// TIA Portal project "OmronFQ2sensor30012026HardInterupt2IRT" (V17)

(* hardware
DEVICE "S7-1200 station_1"  S7-1200 Station
   slot 0: "Rack_0"  S7-1200 Rack  Rack  V1.0
   slot 1: "PLC_1"  CPU 1215C DC/DC/Rly  6ES7 215-1HG40-0XB0  V4.2
DEVICE "FQ2"  GSD.Device.PN
   slot 0: "Rack"  Rack  V1.0
   slot 0: "FQ2"  FQ2-XXX  FQ2-XXX  1.9.0
      slot 0: "FQ2-XXX"  FQ2-XXX  1.9.0
      slot 1: "Interface"  Interface
         slot 1: "Port 1"  Port 1
      slot 1: "Output Data_1"  Output Data  1.9.0
         slot 0: "Output Data"  Output Data  1.9.0
   slot 2: "Results Data - 32 items_1"  Results Data - 32 items  1.9.0
      slot 0: "Results Data - 32 items"  Results Data - 32 items  1.9.0
DEVICE "GSD device_1"  GSD.Device.PN
   slot 0: "Rack"  Rack  V1.0
   slot 0: "FQ22"  FQ2-XXX  FQ2-XXX  1.9.0
      slot 0: "FQ2-XXX"  FQ2-XXX  1.9.0
      slot 1: "Interface"  Interface
         slot 1: "Port 1"  Port 1
      slot 1: "Output Data_1"  Output Data  1.9.0
         slot 0: "Output Data"  Output Data  1.9.0
   slot 2: "Results Data - 32 items_1"  Results Data - 32 items  1.9.0
      slot 0: "Results Data - 32 items"  Results Data - 32 items  1.9.0
*)

// ===== PLC "PLC_1"  CPU 1215C DC/DC/Rly =====

VAR_GLOBAL   // PLC tag table "FQ2"
   "HWCurrentImpulseEncoder" AT %ID1000 : DInt;   // Значение счётчика энкодера в CPU
   "Input_Discret_Sensor_Product" AT %I0.7 : Bool;   // Входа наличия продукта
   "DOPusher" AT %Q0.0 : Bool;   // Выхода на отбраковщик
   "TemplVariable1ForFront" AT %M100.0 : Bool;   // Временая переменная для формирования фронта счёт продука
   "TempleVarible2ForFront" AT %M100.1 : Bool;   // Временая переменая для формирования фронта счёта брака
   "TempleVarible3ForFront" AT %M100.2 : Bool;
   "Tag_1" AT %M100.5 : Bool;
   "Tag_2" AT %M10.1 : Bool;
   "TempleVarible4ForFront" AT %M100.3 : Bool;
   "TempleVarible5ForFront" AT %M100.4 : Bool;
   "Tag_3" AT %M0.0 : Bool;
END_VAR

DATA_BLOCK "QueueProduct_1"   // DB1
{ S7_Optimized_Access := 'FALSE' }
VERSION : 0.1
   VAR
      StructQueue : Array[0..100] of Struct
         QueueAwaitingTrigerCam : Bool;   // Бит ожидания в очереди по камере
         QueueAwaitingRejection : Bool;   // Бит ожидания в очереди по отбраковке
         AwaitingDistanceCamera : Bool;   // Бит ожидание пройденой дистанции до камеры
         ActiveTrigerCam : Bool;   // Бит на измерение камеры
         AwaitingResultatMeasurement : Bool;   // Бит состояния ожидания ответа от камеры
         ResultMeasurementCamera : Bool;   // Результат полученый от камеры 0-ок 1-брак
         ResultRecieved : Bool;   // Результат получен
         RejectionOn : Bool;   // Активент отбраковщик
         CurrentImpulseEncodera : DInt;
      END_STRUCT;
   END_VAR
BEGIN
END_DATA_BLOCK

DATA_BLOCK "InputOutputCamer"   // DB2
{ S7_Optimized_Access := 'FALSE' }
VERSION : 0.1
   VAR
      InputFromCamera1 : Struct
         FLG : Bool;
         BUSY : Bool;
         Ready : Bool;
         "OR" : Bool;
         RUN : Bool;
         Resv : Bool;
         Resv_1 : Bool;
         Resv_2 : Bool;
         Resv_3 : Bool;
         Resv_4 : Bool;
         Resv_5 : Bool;
         Resv_6 : Bool;
         Resv_7 : Bool;
         Resv_8 : Bool;
         Resv_9 : Bool;
         Error : Bool;
         Gate : Bool;
         Resv_10 : Bool;
         Resv_11 : Bool;
         Resv_12 : Bool;
         Resv_13 : Bool;
         Resv_14 : Bool;
         Resv_15 : Bool;
         Resv_16 : Bool;
         Resv_17 : Bool;
         Resv_18 : Bool;
         Resv_19 : Bool;
         Resv_20 : Bool;
         Resv_21 : Bool;
         Resv_22 : Bool;
         Resv_23 : Bool;
         Resv_24 : Bool;
         CommandCode : Array[0..1] of Word;
         ResponseCode : Array[0..3] of Byte;
         ResponseData : Array[0..3] of Byte;
         OutputData1 : Array[0..3] of Byte;
         OutputData2 : Array[0..3] of Byte;
         OutputData3 : Array[0..3] of Byte;
         OutputData4 : Array[0..3] of Byte;
         OutputData5 : Array[0..3] of Byte;
         OutputData6 : Array[0..3] of Byte;
         OutputData7 : Array[0..3] of Byte;
         OutputData8 : Array[0..3] of Byte;
         OutputData9 : Array[0..3] of Byte;
         OutputData10 : Array[0..3] of Byte;
         OutputData11 : Array[0..3] of Byte;
         OutputData12 : Array[0..3] of Byte;
         OutputData13 : Array[0..3] of Byte;
         OutputData14 : Array[0..3] of Byte;
         OutputData15 : Array[0..3] of Byte;
         OutputData16 : Array[0..3] of Byte;
         OutputData17 : Array[0..3] of Byte;
         OutputData18 : Array[0..3] of Byte;
         OutputData19 : Array[0..3] of Byte;
         OutputData20 : Array[0..3] of Byte;
         OutputData21 : Array[0..3] of Byte;
         OutputData22 : Array[0..3] of Byte;
         OutputData23 : Array[0..3] of Byte;
         OutputData24 : Array[0..3] of Byte;
         OutputData25 : Array[0..3] of Byte;
         OutputData26 : Array[0..3] of Byte;
         OutputData27 : Array[0..3] of Byte;
         OutputData28 : Array[0..3] of Byte;
         OutputData29 : Array[0..3] of Byte;
         OutputData30 : Array[0..3] of Byte;
         OutputData31 : Array[0..3] of Byte;
         OutputData32 : Array[0..3] of Byte;
      END_STRUCT;
      OutputFromPLCtoCamera1 : Struct
         EXE : Bool;
         TRIG : Bool;
         Resv : Bool;
         Resv_1 : Bool;
         Resv_2 : Bool;
         Resv_3 : Bool;
         Resv_4 : Bool;
         Resv_5 : Bool;
         Resv_6 : Bool;
         Resv_7 : Bool;
         Resv_8 : Bool;
         Resv_9 : Bool;
         Resv_10 : Bool;
         Resv_11 : Bool;
         Resv_12 : Bool;
         ERCLR : Bool;
         DSA : Bool;
         Resv_13 : Bool;
         Resv_14 : Bool;
         Resv_15 : Bool;
         Resv_16 : Bool;
         Resv_17 : Bool;
         Resv_18 : Bool;
         Resv_19 : Bool;
         Resv_20 : Bool;
         Resv_21 : Bool;
         Resv_22 : Bool;
         Resv_23 : Bool;
         Resv_24 : Bool;
         Resv_25 : Bool;
         Resv_26 : Bool;
         Resv_27 : Bool;
         ComandCode : Array[0..1] of Word;
         ComandParameter : Array[0..3] of Byte;
         ComandParameter2 : Array[0..3] of Byte;
         ComandParameter3 : Array[0..3] of Byte;
      END_STRUCT;
      InputFromCamera2 : Struct
         FLG : Bool;
         BUSY : Bool;
         Ready : Bool;
         "OR" : Bool;
         RUN : Bool;
         Resv : Bool;
         Resv_1 : Bool;
         Resv_2 : Bool;
         Resv_3 : Bool;
         Resv_4 : Bool;
         Resv_5 : Bool;
         Resv_6 : Bool;
         Resv_7 : Bool;
         Resv_8 : Bool;
         Resv_9 : Bool;
         Error : Bool;
         Gate : Bool;
         Resv_10 : Bool;
         Resv_11 : Bool;
         Resv_12 : Bool;
         Resv_13 : Bool;
         Resv_14 : Bool;
         Resv_15 : Bool;
         Resv_16 : Bool;
         Resv_17 : Bool;
         Resv_18 : Bool;
         Resv_19 : Bool;
         Resv_20 : Bool;
         Resv_21 : Bool;
         Resv_22 : Bool;
         Resv_23 : Bool;
         Resv_24 : Bool;
         CommandCode : Array[0..1] of Word;
         ResponseCode : Array[0..3] of Byte;
         ResponseData : Array[0..3] of Byte;
         OutputData1 : Array[0..3] of Byte;
         OutputData2 : Array[0..3] of Byte;
         OutputData3 : Array[0..3] of Byte;
         OutputData4 : Array[0..3] of Byte;
         OutputData5 : Array[0..3] of Byte;
         OutputData6 : Array[0..3] of Byte;
         OutputData7 : Array[0..3] of Byte;
         OutputData8 : Array[0..3] of Byte;
         OutputData9 : Array[0..3] of Byte;
         OutputData10 : Array[0..3] of Byte;
         OutputData11 : Array[0..3] of Byte;
         OutputData12 : Array[0..3] of Byte;
         OutputData13 : Array[0..3] of Byte;
         OutputData14 : Array[0..3] of Byte;
         OutputData15 : Array[0..3] of Byte;
         OutputData16 : Array[0..3] of Byte;
         OutputData17 : Array[0..3] of Byte;
         OutputData18 : Array[0..3] of Byte;
         OutputData19 : Array[0..3] of Byte;
         OutputData20 : Array[0..3] of Byte;
         OutputData21 : Array[0..3] of Byte;
         OutputData22 : Array[0..3] of Byte;
         OutputData23 : Array[0..3] of Byte;
         OutputData24 : Array[0..3] of Byte;
         OutputData25 : Array[0..3] of Byte;
         OutputData26 : Array[0..3] of Byte;
         OutputData27 : Array[0..3] of Byte;
         OutputData28 : Array[0..3] of Byte;
         OutputData29 : Array[0..3] of Byte;
         OutputData30 : Array[0..3] of Byte;
         OutputData31 : Array[0..3] of Byte;
         OutputData32 : Array[0..3] of Byte;
      END_STRUCT;
      OutputFromPLCtoCamera2 : Struct
         EXE : Bool;
         TRIG : Bool;
         Resv : Bool;
         Resv_1 : Bool;
         Resv_2 : Bool;
         Resv_3 : Bool;
         Resv_4 : Bool;
         Resv_5 : Bool;
         Resv_6 : Bool;
         Resv_7 : Bool;
         Resv_8 : Bool;
         Resv_9 : Bool;
         Resv_10 : Bool;
         Resv_11 : Bool;
         Resv_12 : Bool;
         ERCLR : Bool;
         DSA : Bool;
         Resv_13 : Bool;
         Resv_14 : Bool;
         Resv_15 : Bool;
         Resv_16 : Bool;
         Resv_17 : Bool;
         Resv_18 : Bool;
         Resv_19 : Bool;
         Resv_20 : Bool;
         Resv_21 : Bool;
         Resv_22 : Bool;
         Resv_23 : Bool;
         Resv_24 : Bool;
         Resv_25 : Bool;
         Resv_26 : Bool;
         Resv_27 : Bool;
         ComandCode : Array[0..1] of Word;
         ComandParameter : Array[0..3] of Byte;
         ComandParameter2 : Array[0..3] of Byte;
         ComandParameter3 : Array[0..3] of Byte;
      END_STRUCT;
   END_VAR
BEGIN
   InputFromCamera1.CommandCode[0] := 16#0;
   InputFromCamera2.CommandCode[0] := 16#0;
END_DATA_BLOCK

DATA_BLOCK "AuxaluryBlockProcesseComandeCamera"   // DB3
{ S7_Optimized_Access := 'FALSE' }
VERSION : 0.1
   VAR
      RequestComandeFromPlcToCamera_1 : Bool;   // Бит начала запроса выполнения команды с плк на камеру
      RequestConfirmComandeFromPLCtoCamera_1 : Bool;   // Бит подтверждения что запрос команды отправлен
      RequestComandeFromPlcToCamera_2 : Bool;
      RequestConfirmComandeFromPLCtoCamera_2 : Bool;
      Camera1ChangeSceneOk : Bool;
      Camera2ChangeSceneOk : Bool;
      QuitRejectCam1 : Bool;   // Отбраковка по камере 1
      QuitRejectCam2 : Bool;   // Отбраковка по камере 2
      RequestChangeSceneCamera1 : Bool;   // Дополнительный бить для обработки переключения рецецтпа камеры 1
      RequestChangeSceneCamera2 : Bool;   // Дополнительный бить для обработки переключения рецецтпа камеры 2
   END_VAR
BEGIN
END_DATA_BLOCK

DATA_BLOCK "QueueProduct_2"   // DB4
{ S7_Optimized_Access := 'TRUE' }
VERSION : 0.1
   VAR
      StructQueue : Array[0..100] of Struct
         QueueAwaitingTrigerCam : Bool;   // Бит ожидания в очереди по камере
         QueueAwaitingRejection : Bool;   // Бит ожидания в очереди по отбраковке
         AwaitingDistanceCamera : Bool;   // Бит ожидание пройденой дистанции до камеры
         ActiveTrigerCam : Bool;   // Бит на измерение камеры
         AwaitingResultatMeasurement : Bool;   // Бит состояния ожидания ответа от камеры
         ResultMeasurementCamera : Bool;   // Результат полученый от камеры 0-ок 1-брак
         ResultRecieved : Bool;   // Результат получен
         RejectionOn : Bool;   // Активент отбраковщик
         CurrentImpulseEncodera : DInt;
      END_STRUCT;
   END_VAR
BEGIN
END_DATA_BLOCK

DATA_BLOCK "DataBlockHMI"   // DB5
{ S7_Optimized_Access := 'FALSE' }
VERSION : 0.1
   VAR
      CountProduct : UDInt;   // Кол-во продукта прошедшего отбраковщик
      CountRejection : UDInt;   // Кол-во отбракованного
      NumberSceneRequest : Byte;   // Запрос номера сценария в камере
      Buttons : Struct
         ButtonChangeRecipe : Bool;   // Кнопка запрос на изменение рецепта(сцены)камеры от оператора
         ButtonWorkRestrictionPusher : Bool;   // Кнопка запрета работы пушера отбраковщика
         ButtonLoadFromActualInList : Bool;
         ButtonWorkOffCam1 : Bool;   // Камера 1 не обрабатывает очередь продукта
         ButtonWorkOffCam2 : Bool;   // Камера 2 не обрабатывает очередь продукта
         Button5 : Bool;
         Button6 : Bool;
         Button7 : Bool;
      END_STRUCT;
      AuxilaryBit : Array[0..7] of Bool;
      Recipe : Array[0..32] of Struct
         CountImpTrigerCamera1 : DInt;   // Количество импульсов для сработки камеры
         CountImpForRegection1 : DInt;   // Количество импульсов для отбраковки
         CountImpForResetRegectio1 : DInt;   // Количество импульсов для длительности отбраковки
         NumberRecipeScene : Byte;   // Номер сценария в камере
         HighMM : Int;   // высота в милиметрах
         OverhangValue : Int;   // величина вылета в милиметрах
         CountImpTrigerCamera2 : DInt;
         CountImpForRegection2 : DInt;
      END_STRUCT;
      CountRejectionCam1 : UDInt;   // Количество отбраковоаного по камере 1
      CountRejectionCam2 : UDInt;   // Количество отбракованого по камере 2
   END_VAR
BEGIN
   Recipe[0].CountImpTrigerCamera1 := 335;
   Recipe[0].CountImpForRegection1 := 455;
   Recipe[0].CountImpForResetRegectio1 := 25;
   Recipe[0].NumberRecipeScene := 0;
   Recipe[1].CountImpTrigerCamera1 := 335;
   Recipe[1].CountImpForRegection1 := 455;
   Recipe[1].CountImpForResetRegectio1 := 25;
   Recipe[1].NumberRecipeScene := 0;
   Recipe[2].CountImpTrigerCamera1 := 335;
   Recipe[2].CountImpForRegection1 := 455;
   Recipe[2].CountImpForResetRegectio1 := 25;
   Recipe[2].NumberRecipeScene := 1;
   Recipe[3].CountImpTrigerCamera1 := 335;
   Recipe[3].CountImpForRegection1 := 455;
   Recipe[3].CountImpForResetRegectio1 := 25;
   Recipe[3].NumberRecipeScene := 2;
   Recipe[4].CountImpTrigerCamera1 := 335;
   Recipe[4].CountImpForRegection1 := 455;
   Recipe[4].CountImpForResetRegectio1 := 25;
   Recipe[4].NumberRecipeScene := 3;
   Recipe[5].CountImpTrigerCamera1 := 335;
   Recipe[5].CountImpForRegection1 := 455;
   Recipe[5].CountImpForResetRegectio1 := 25;
   Recipe[5].NumberRecipeScene := 4;
   Recipe[6].CountImpTrigerCamera1 := 335;
   Recipe[6].CountImpForRegection1 := 455;
   Recipe[6].CountImpForResetRegectio1 := 25;
   Recipe[6].NumberRecipeScene := 5;
   Recipe[7].CountImpTrigerCamera1 := 335;
   Recipe[7].CountImpForRegection1 := 455;
   Recipe[7].CountImpForResetRegectio1 := 25;
   Recipe[7].NumberRecipeScene := 6;
   Recipe[8].CountImpTrigerCamera1 := 335;
   Recipe[8].CountImpForRegection1 := 455;
   Recipe[8].CountImpForResetRegectio1 := 25;
   Recipe[8].NumberRecipeScene := 7;
   Recipe[9].CountImpTrigerCamera1 := 335;
   Recipe[9].CountImpForRegection1 := 455;
   Recipe[9].CountImpForResetRegectio1 := 25;
   Recipe[9].NumberRecipeScene := 8;
   Recipe[10].CountImpTrigerCamera1 := 335;
   Recipe[10].CountImpForRegection1 := 455;
   Recipe[10].CountImpForResetRegectio1 := 25;
   Recipe[10].NumberRecipeScene := 9;
   Recipe[11].CountImpTrigerCamera1 := 335;
   Recipe[11].CountImpForRegection1 := 455;
   Recipe[11].CountImpForResetRegectio1 := 25;
   Recipe[11].NumberRecipeScene := 10;
   Recipe[12].CountImpTrigerCamera1 := 335;
   Recipe[12].CountImpForRegection1 := 455;
   Recipe[12].CountImpForResetRegectio1 := 25;
   Recipe[12].NumberRecipeScene := 11;
   Recipe[13].CountImpTrigerCamera1 := 335;
   Recipe[13].CountImpForRegection1 := 455;
   Recipe[13].CountImpForResetRegectio1 := 25;
   Recipe[13].NumberRecipeScene := 12;
   Recipe[14].CountImpTrigerCamera1 := 335;
   Recipe[14].CountImpForRegection1 := 455;
   Recipe[14].CountImpForResetRegectio1 := 25;
   Recipe[14].NumberRecipeScene := 13;
   Recipe[15].CountImpTrigerCamera1 := 335;
   Recipe[15].CountImpForRegection1 := 455;
   Recipe[15].CountImpForResetRegectio1 := 25;
   Recipe[15].NumberRecipeScene := 14;
   Recipe[16].CountImpTrigerCamera1 := 335;
   Recipe[16].CountImpForRegection1 := 455;
   Recipe[16].CountImpForResetRegectio1 := 25;
   Recipe[16].NumberRecipeScene := 15;
   Recipe[17].CountImpTrigerCamera1 := 335;
   Recipe[17].CountImpForRegection1 := 455;
   Recipe[17].CountImpForResetRegectio1 := 25;
   Recipe[17].NumberRecipeScene := 16;
   Recipe[18].CountImpTrigerCamera1 := 335;
   Recipe[18].CountImpForRegection1 := 455;
   Recipe[18].CountImpForResetRegectio1 := 25;
   Recipe[18].NumberRecipeScene := 17;
   Recipe[19].CountImpTrigerCamera1 := 335;
   Recipe[19].CountImpForRegection1 := 455;
   Recipe[19].CountImpForResetRegectio1 := 25;
   Recipe[19].NumberRecipeScene := 18;
   Recipe[20].CountImpTrigerCamera1 := 335;
   Recipe[20].CountImpForRegection1 := 455;
   Recipe[20].CountImpForResetRegectio1 := 25;
   Recipe[20].NumberRecipeScene := 19;
   Recipe[21].CountImpTrigerCamera1 := 335;
   Recipe[21].CountImpForRegection1 := 455;
   Recipe[21].CountImpForResetRegectio1 := 25;
   Recipe[21].NumberRecipeScene := 20;
   Recipe[22].CountImpTrigerCamera1 := 335;
   Recipe[22].CountImpForRegection1 := 455;
   Recipe[22].CountImpForResetRegectio1 := 25;
   Recipe[22].NumberRecipeScene := 21;
   Recipe[23].CountImpTrigerCamera1 := 335;
   Recipe[23].CountImpForRegection1 := 455;
   Recipe[23].CountImpForResetRegectio1 := 25;
   Recipe[23].NumberRecipeScene := 22;
   Recipe[24].CountImpTrigerCamera1 := 335;
   Recipe[24].CountImpForRegection1 := 455;
   Recipe[24].CountImpForResetRegectio1 := 25;
   Recipe[24].NumberRecipeScene := 23;
   Recipe[25].CountImpTrigerCamera1 := 335;
   Recipe[25].CountImpForRegection1 := 455;
   Recipe[25].CountImpForResetRegectio1 := 25;
   Recipe[25].NumberRecipeScene := 24;
   Recipe[26].CountImpTrigerCamera1 := 335;
   Recipe[26].CountImpForRegection1 := 455;
   Recipe[26].CountImpForResetRegectio1 := 25;
   Recipe[26].NumberRecipeScene := 25;
   Recipe[27].CountImpTrigerCamera1 := 335;
   Recipe[27].CountImpForRegection1 := 455;
   Recipe[27].CountImpForResetRegectio1 := 25;
   Recipe[27].NumberRecipeScene := 26;
   Recipe[28].CountImpTrigerCamera1 := 335;
   Recipe[28].CountImpForRegection1 := 455;
   Recipe[28].CountImpForResetRegectio1 := 25;
   Recipe[28].NumberRecipeScene := 27;
   Recipe[29].CountImpTrigerCamera1 := 335;
   Recipe[29].CountImpForRegection1 := 455;
   Recipe[29].CountImpForResetRegectio1 := 25;
   Recipe[29].NumberRecipeScene := 28;
   Recipe[30].CountImpTrigerCamera1 := 335;
   Recipe[30].CountImpForRegection1 := 455;
   Recipe[30].CountImpForResetRegectio1 := 25;
   Recipe[30].NumberRecipeScene := 29;
   Recipe[31].CountImpTrigerCamera1 := 335;
   Recipe[31].CountImpForRegection1 := 455;
   Recipe[31].CountImpForResetRegectio1 := 25;
   Recipe[31].NumberRecipeScene := 30;
   Recipe[32].CountImpTrigerCamera1 := 335;
   Recipe[32].CountImpForRegection1 := 455;
   Recipe[32].CountImpForResetRegectio1 := 25;
   Recipe[32].NumberRecipeScene := 31;
   // AuxilaryBit[0] : Бит для подсчёта брака cam1
   // Recipe[0] : Действующей рецепт(сценарий)
   // Recipe[1] : Сценарий 0
   // Recipe[2] : Сценарий 1
   // Recipe[3] : Сценарий 2
   // Recipe[4] : Сценарий 3
   // Recipe[5] : Сценарий 4
   // Recipe[6] : Сценарий 5
   // Recipe[7] : Сценарий 6
   // Recipe[8] : Сценарий 7
   // Recipe[9] : Сценарий 8
   // Recipe[10] : Сценарий 9
   // AuxilaryBit[1] : Бит для подсчёта брака сam2
END_DATA_BLOCK

FUNCTION "QueueCreate" : Void   // FC3, SCL
{ S7_Optimized_Access := 'FALSE' }
VERSION : 0.1
   VAR_TEMP
      i1 : Int;
      i2 : Int;
      d : Int;
   END_VAR
BEGIN
   //Добовляем в очередь продукт

       FOR #i1 := 0 TO 20 DO
           // Statement section FOR
           IF NOT "QueueProduct_1".StructQueue[#i1].QueueAwaitingRejection THEN
               IF NOT "DataBlockHMI".Buttons.ButtonWorkOffCam1 THEN //условие чтоб камеру выключить не обрабоатывать ничего
                   "QueueProduct_1".StructQueue[#i1].QueueAwaitingTrigerCam := TRUE;
                   "QueueProduct_1".StructQueue[#i1].QueueAwaitingRejection := TRUE;
               END_IF;

               EXIT;
           END_IF;
       END_FOR;
       FOR #i2 := 0 TO 20 DO
           // Statement section FOR
           IF NOT "QueueProduct_2".StructQueue[#i2].QueueAwaitingRejection THEN
               IF NOT "DataBlockHMI".Buttons.ButtonWorkOffCam2 THEN
                   "QueueProduct_2".StructQueue[#i2].QueueAwaitingTrigerCam := TRUE;
                   "QueueProduct_2".StructQueue[#i2].QueueAwaitingRejection := TRUE;
               END_IF;
               EXIT;
           END_IF;
       END_FOR;

   "DataBlockHMI".CountProduct := UDINT#1 + "DataBlockHMI".CountProduct;

   IF NOT "DataBlockHMI".Buttons.ButtonWorkOffCam1 THEN
       "ProcessingQueue1"(NumberQueue := #i1); //Обрабатываем только что добавленую очередь
   END_IF;
   IF NOT "DataBlockHMI".Buttons.ButtonWorkOffCam2 THEN
       "ProcessingQueue2"(NumberQueue := #i2);
   END_IF;
END_FUNCTION

FUNCTION "ProcessingQueue1" : Void   // FC4, SCL
{ S7_Optimized_Access := 'TRUE' }
VERSION : 0.1
   VAR_INPUT
      NumberQueue : Int;
   END_VAR
BEGIN
   IF  "QueueProduct_1".StructQueue[#NumberQueue].QueueAwaitingRejection THEN
       // Statement section IF


       //Создание запроса в очереди на тригер камеры, запоминаем текущие положение продукта
       IF "QueueProduct_1".StructQueue[#NumberQueue].QueueAwaitingTrigerCam &
           "QueueProduct_1".StructQueue[#NumberQueue].QueueAwaitingRejection THEN

           "QueueProduct_1".StructQueue[#NumberQueue].CurrentImpulseEncodera := "HWCurrentImpulseEncoder":P;
           "QueueProduct_1".StructQueue[#NumberQueue].QueueAwaitingTrigerCam := False;
           "QueueProduct_1".StructQueue[#NumberQueue].AwaitingDistanceCamera := True;
           RETURN;
       END_IF;
       //Выходим из проверки пока продукт не доехал до камеры, оптимизация чтоб не пробегать всю функцию
       IF "QueueProduct_1".StructQueue[#NumberQueue].CurrentImpulseEncodera +"DataBlockHMI".Recipe[0].CountImpTrigerCamera1(*Recip[0] прният как действующей рецепт*) >"HWCurrentImpulseEncoder":P THEN
           RETURN;
       END_IF;    
           //По прохождению дистанции взводим бит для работы камеры, снимаем бит ожидания 
       IF "QueueProduct_1".StructQueue[#NumberQueue].AwaitingDistanceCamera
           &"QueueProduct_1".StructQueue[#NumberQueue].CurrentImpulseEncodera + "DataBlockHMI".Recipe[0].CountImpTrigerCamera1(*Recip[0] прният как действующей рецепт*) <="HWCurrentImpulseEncoder":P
            & NOT "InputOutputCamer".InputFromCamera1.BUSY THEN

           "QueueProduct_1".StructQueue[#NumberQueue].ActiveTrigerCam := true;
           "InputOutputCamer".OutputFromPLCtoCamera1.TRIG := true;
           "QueueProduct_1".StructQueue[#NumberQueue].AwaitingDistanceCamera := False;
           RETURN;
       END_IF;

       //На период обработки камеры снимаем бит работы камеры, взводим бит ожидание ответа от камеры
       IF "QueueProduct_1".StructQueue[#NumberQueue].ActiveTrigerCam & "InputOutputCamer".InputFromCamera1.BUSY THEN

           "QueueProduct_1".StructQueue[#NumberQueue].ActiveTrigerCam := False;
           "InputOutputCamer".OutputFromPLCtoCamera1.TRIG := false;
           "QueueProduct_1".StructQueue[#NumberQueue].AwaitingResultatMeasurement := True;
           RETURN;
       END_IF;

       //Ожидание получение ответа от камеры, фиксируем что ответ был
       IF "QueueProduct_1".StructQueue[#NumberQueue].AwaitingResultatMeasurement & NOT "InputOutputCamer".InputFromCamera1.BUSY
       THEN

           "QueueProduct_1".StructQueue[#NumberQueue].ResultMeasurementCamera := "InputOutputCamer".InputFromCamera1."OR";
           "QueueProduct_1".StructQueue[#NumberQueue].ResultRecieved := True;
           "QueueProduct_1".StructQueue[#NumberQueue].AwaitingResultatMeasurement := FALSE;

       END_IF;

       //Обработка полученого ответа от камеры(бракуем или нет).
       //Если не бракуем, освобождаем очередь, Если бракуем то взводим бит браковки и освобождаем очередь после снятия сигнала с пушера
       IF "QueueProduct_1".StructQueue[#NumberQueue].ResultRecieved & "QueueProduct_1".StructQueue[#NumberQueue].ResultMeasurementCamera
           & ("QueueProduct_1".StructQueue[#NumberQueue].CurrentImpulseEncodera + "DataBlockHMI".Recipe[0].CountImpTrigerCamera1
           + "DataBlockHMI".Recipe[0].CountImpForRegection1 <= "HWCurrentImpulseEncoder":P) THEN //условия для старта отбраковки

           "AuxaluryBlockProcesseComandeCamera".QuitRejectCam1 := true;
           "DataBlockHMI".AuxilaryBit[0] := TRUE;
           "QueueProduct_1".StructQueue[#NumberQueue].RejectionOn := true;
           "QueueProduct_1".StructQueue[#NumberQueue].ResultRecieved := FALSE;

       ELSIF "QueueProduct_1".StructQueue[#NumberQueue].ResultRecieved & NOT "QueueProduct_1".StructQueue[#NumberQueue].ResultMeasurementCamera THEN

           "QueueProduct_1".StructQueue[#NumberQueue] := "QueueProduct_1".StructQueue[100];

       END_IF;

       //Cнимаем выход отбраковки и скидываем очередь
       IF "QueueProduct_1".StructQueue[#NumberQueue].RejectionOn & ("QueueProduct_1".StructQueue[#NumberQueue].CurrentImpulseEncodera + "DataBlockHMI".Recipe[0].CountImpTrigerCamera1
           + "DataBlockHMI".Recipe[0].CountImpForRegection1 +"DataBlockHMI".Recipe[0].CountImpForResetRegectio1 <="HWCurrentImpulseEncoder":P) THEN

           "AuxaluryBlockProcesseComandeCamera".QuitRejectCam1 := false;
           "DataBlockHMI".AuxilaryBit[0] := FALSE;
           "QueueProduct_1".StructQueue[#NumberQueue] := "QueueProduct_1".StructQueue[100];

       END_IF;

       IF "DataBlockHMI".Buttons.ButtonWorkRestrictionPusher THEN
           "AuxaluryBlockProcesseComandeCamera".QuitRejectCam1 := FALSE;

       END_IF;


   END_IF;
END_FUNCTION

FUNCTION "ChangeSceneOnCameraFQ2" : Void   // FC6, SCL
{ S7_Optimized_Access := 'FALSE' }
VERSION : 0.1
   VAR_INPUT
      NumberScene : Byte;
   END_VAR
   VAR_IN_OUT
      RequestChangeScene : Bool;
   END_VAR
BEGIN
   //Запроc смены рецепта или есть ожидание от прошлого выполняем
   //условия обработки смены сценария, здесь создаём защиту от зацикливания
   //посредсвом проверки прошлый запрос прошёл успешно и ждём вторую камеру

   IF #RequestChangeScene AND NOT "AuxaluryBlockProcesseComandeCamera".RequestChangeSceneCamera1 AND NOT "AuxaluryBlockProcesseComandeCamera".Camera1ChangeSceneOk THEN
          "AuxaluryBlockProcesseComandeCamera".RequestChangeSceneCamera1 := TRUE;
      END_IF;

   IF #RequestChangeScene AND NOT "AuxaluryBlockProcesseComandeCamera".RequestChangeSceneCamera2 AND NOT "AuxaluryBlockProcesseComandeCamera".Camera2ChangeSceneOk THEN
         "AuxaluryBlockProcesseComandeCamera".RequestChangeSceneCamera2 := TRUE;
   END_IF;


   // Команда на камеру1 для выполнения переключения сценария проверки и номер сценария
      IF "AuxaluryBlockProcesseComandeCamera".RequestChangeSceneCamera1 AND NOT "InputOutputCamer".InputFromCamera1.BUSY
          AND NOT "AuxaluryBlockProcesseComandeCamera".Camera1ChangeSceneOk THEN


         "InputOutputCamer".OutputFromPLCtoCamera1.ComandCode[0] := 16#30;
         "InputOutputCamer".OutputFromPLCtoCamera1.ComandCode[1] := 16#1000;
         "InputOutputCamer".OutputFromPLCtoCamera1.ComandParameter[3] := #NumberScene;
         "AuxaluryBlockProcesseComandeCamera".RequestConfirmComandeFromPLCtoCamera_1 := TRUE;
         "InputOutputCamer".OutputFromPLCtoCamera1.EXE := TRUE;

     END_IF;

   // Команда на камеру2 для выполнения переключения сценария проверки и номер сценария
     IF "AuxaluryBlockProcesseComandeCamera".RequestChangeSceneCamera2 AND NOT "InputOutputCamer".InputFromCamera2.BUSY
         AND NOT "AuxaluryBlockProcesseComandeCamera".Camera2ChangeSceneOk THEN


         "InputOutputCamer".OutputFromPLCtoCamera2.ComandCode[0] := 16#30;
         "InputOutputCamer".OutputFromPLCtoCamera2.ComandCode[1] := 16#1000;
         "InputOutputCamer".OutputFromPLCtoCamera2.ComandParameter[3] := #NumberScene;
         "AuxaluryBlockProcesseComandeCamera".RequestConfirmComandeFromPLCtoCamera_2 := TRUE;
         "InputOutputCamer".OutputFromPLCtoCamera2.EXE := TRUE;

     END_IF;

       // После послания запроса ожидаем возвращени выполнения подтверждения от камеры 1, что всё выполнено и сбрасываем биты и команды.
     IF "AuxaluryBlockProcesseComandeCamera".RequestConfirmComandeFromPLCtoCamera_1
         AND "InputOutputCamer".InputFromCamera1.BUSY
         AND "InputOutputCamer".InputFromCamera1.FLG AND NOT "AuxaluryBlockProcesseComandeCamera".Camera1ChangeSceneOk THEN

         //#RequestChangeScene := FALSE;
         "AuxaluryBlockProcesseComandeCamera".RequestConfirmComandeFromPLCtoCamera_1 := FALSE;
         "InputOutputCamer".OutputFromPLCtoCamera1.EXE := False;
         "InputOutputCamer".OutputFromPLCtoCamera1.ComandCode[0] := 16#0;
         "InputOutputCamer".OutputFromPLCtoCamera1.ComandCode[1] := 16#0;
         "InputOutputCamer".OutputFromPLCtoCamera1.ComandParameter[3] := 0;
         IF "InputOutputCamer".InputFromCamera1.ResponseCode[0] = 0
             AND
             "InputOutputCamer".InputFromCamera1.ResponseCode[1] = 0
             AND
             "InputOutputCamer".InputFromCamera1.ResponseCode[2] = 0
             AND
             "InputOutputCamer".InputFromCamera1.ResponseCode[3] = 0
         THEN
             "AuxaluryBlockProcesseComandeCamera".Camera1ChangeSceneOk := TRUE;
         END_IF;
         //#RequestChangeScene := False;
     END_IF;

    // После послания запроса ожидаем возвращени выполнения подтверждения от камеры 2, что всё выполнено и сбрасываем биты и команды.
     IF "AuxaluryBlockProcesseComandeCamera".RequestConfirmComandeFromPLCtoCamera_2
         AND "InputOutputCamer".InputFromCamera2.BUSY
         AND "InputOutputCamer".InputFromCamera2.FLG AND NOT "AuxaluryBlockProcesseComandeCamera".Camera2ChangeSceneOk THEN

         //#RequestChangeScene := FALSE;
         "AuxaluryBlockProcesseComandeCamera".RequestConfirmComandeFromPLCtoCamera_2 := FALSE;
         "InputOutputCamer".OutputFromPLCtoCamera2.EXE := False;
         "InputOutputCamer".OutputFromPLCtoCamera2.ComandCode[0] := 16#0;
         "InputOutputCamer".OutputFromPLCtoCamera2.ComandCode[1] := 16#0;
         "InputOutputCamer".OutputFromPLCtoCamera2.ComandParameter[3] := 0;
         IF "InputOutputCamer".InputFromCamera2.ResponseCode[0] = 0
             AND
             "InputOutputCamer".InputFromCamera2.ResponseCode[1] = 0
             AND
             "InputOutputCamer".InputFromCamera2.ResponseCode[2] = 0
             AND
             "InputOutputCamer".InputFromCamera2.ResponseCode[3] = 0
         THEN
             "AuxaluryBlockProcesseComandeCamera".Camera2ChangeSceneOk:=TRUE;
         END_IF;
         //#RequestChangeScene := False;
     END_IF;
     (* IF "AuxaluryBlockProcesseComandeCamera".Camera1ChangeSceneOk  THEN
         "RecipeFromListToActual"(#NumberScene);
         //"AuxaluryBlockProcesseComandeCamera".Camera2ChangeSceneOk := FALSE;
         "AuxaluryBlockProcesseComandeCamera".Camera1ChangeSceneOk := FALSE;

     END_IF;

     IF "AuxaluryBlockProcesseComandeCamera".Camera2ChangeSceneOk THEN
         "RecipeFromListToActual"(#NumberScene);
         "AuxaluryBlockProcesseComandeCamera".Camera2ChangeSceneOk := FALSE;
         //"AuxaluryBlockProcesseComandeCamera".Camera1ChangeSceneOk := FALSE;

     END_IF; *)
     //Cнимаеме повторение запросов
     IF "AuxaluryBlockProcesseComandeCamera".Camera1ChangeSceneOk AND "AuxaluryBlockProcesseComandeCamera".RequestChangeSceneCamera1 THEN

         "AuxaluryBlockProcesseComandeCamera".RequestChangeSceneCamera1 := FALSE;

     END_IF;

     IF "AuxaluryBlockProcesseComandeCamera".Camera2ChangeSceneOk AND "AuxaluryBlockProcesseComandeCamera".RequestChangeSceneCamera2 THEN
         "AuxaluryBlockProcesseComandeCamera".RequestChangeSceneCamera1 := FALSE;
     END_IF;

     //Перенос рецепта из памяти в актуальный работающий сброс битов
     IF "AuxaluryBlockProcesseComandeCamera".Camera1ChangeSceneOk AND "AuxaluryBlockProcesseComandeCamera".Camera2ChangeSceneOk THEN
         "RecipeFromListToActual"(#NumberScene);
         "AuxaluryBlockProcesseComandeCamera".Camera1ChangeSceneOk := FALSE;
         "AuxaluryBlockProcesseComandeCamera".Camera2ChangeSceneOk := FALSE;
         #RequestChangeScene := FALSE;

     END_IF;
END_FUNCTION

FUNCTION "RecipeFromListToActual" : Void   // FC7, SCL
{ S7_Optimized_Access := 'TRUE' }
VERSION : 0.1
   VAR_INPUT
      InputNumber : Byte;   // Указание какой рецепт загружаем в актуальный
   END_VAR
   VAR_TEMP
      i : Int;   // временая переменая для прогона
   END_VAR
BEGIN

   FOR  #i:= 1 TO 32 DO

       IF "DataBlockHMI".Recipe[#i].NumberRecipeScene = #InputNumber THEN

           "DataBlockHMI".Recipe[0] := "DataBlockHMI".Recipe[#i];
           EXIT;
       END_IF;


       END_FOR;
END_FUNCTION

FUNCTION "RecipFromActualToList" : Void   // FC8, SCL
{ S7_Optimized_Access := 'TRUE' }
VERSION : 0.1
   VAR_INPUT
      InputNumber : Byte;
   END_VAR
   VAR_TEMP
      i : Int;
   END_VAR
BEGIN
   FOR #i := 1 TO 32 DO

       IF "DataBlockHMI".Recipe[#i].NumberRecipeScene = #InputNumber THEN

           "DataBlockHMI".Recipe[#i] := "DataBlockHMI".Recipe[0];
           EXIT;
       END_IF;


   END_FOR;
END_FUNCTION

FUNCTION "ProcessingQueue2" : Void   // FC9, SCL
{ S7_Optimized_Access := 'TRUE' }
VERSION : 0.1
   VAR_INPUT
      NumberQueue : Int;
   END_VAR
BEGIN
   IF "QueueProduct_2".StructQueue[#NumberQueue].QueueAwaitingRejection THEN
       // Statement section IF


       //Создание запроса в очереди на тригер камеры, запоминаем текущие положение продукта
       IF "QueueProduct_2".StructQueue[#NumberQueue].QueueAwaitingTrigerCam &
           "QueueProduct_2".StructQueue[#NumberQueue].QueueAwaitingRejection THEN

           "QueueProduct_2".StructQueue[#NumberQueue].CurrentImpulseEncodera := "HWCurrentImpulseEncoder":P;
           "QueueProduct_2".StructQueue[#NumberQueue].QueueAwaitingTrigerCam := False;
           "QueueProduct_2".StructQueue[#NumberQueue].AwaitingDistanceCamera := True;
           RETURN;
       END_IF;
       //Выходим из проверки пока продукт не доехал до камеры, оптимизация чтоб не пробегать всю функцию
       IF "QueueProduct_2".StructQueue[#NumberQueue].CurrentImpulseEncodera + "DataBlockHMI".Recipe[0].CountImpTrigerCamera2 > "HWCurrentImpulseEncoder":P THEN
           RETURN;
       END_IF;
       //По прохождению дистанции взводим бит для работы камеры, снимаем бит ожидания 
       IF  "QueueProduct_2".StructQueue[#NumberQueue].AwaitingDistanceCamera
           & "QueueProduct_2".StructQueue[#NumberQueue].CurrentImpulseEncodera + "DataBlockHMI".Recipe[0].CountImpTrigerCamera2<= "HWCurrentImpulseEncoder":P
           &  NOT "InputOutputCamer".InputFromCamera2.BUSY THEN

           "QueueProduct_2".StructQueue[#NumberQueue].ActiveTrigerCam := true;
           "InputOutputCamer".OutputFromPLCtoCamera2.TRIG := true;
           "QueueProduct_2".StructQueue[#NumberQueue].AwaitingDistanceCamera := False;
           RETURN;
       END_IF;

       //На период обработки камеры снимаем бит работы камеры, взводим бит ожидание ответа от камеры
       IF "QueueProduct_2".StructQueue[#NumberQueue].ActiveTrigerCam & "InputOutputCamer".InputFromCamera2.BUSY THEN

           "QueueProduct_2".StructQueue[#NumberQueue].ActiveTrigerCam := False;
           "InputOutputCamer".OutputFromPLCtoCamera2.TRIG := false;
           "QueueProduct_2".StructQueue[#NumberQueue].AwaitingResultatMeasurement := True;
           RETURN;
       END_IF;

       //Ожидание получение ответа от камеры, фиксируем что ответ был
       IF "QueueProduct_2".StructQueue[#NumberQueue].AwaitingResultatMeasurement & NOT "InputOutputCamer".InputFromCamera2.BUSY
       THEN

           "QueueProduct_2".StructQueue[#NumberQueue].ResultMeasurementCamera := "InputOutputCamer".InputFromCamera2."OR";
           "QueueProduct_2".StructQueue[#NumberQueue].ResultRecieved := True;
           "QueueProduct_2".StructQueue[#NumberQueue].AwaitingResultatMeasurement := FALSE;


       END_IF;

       //Обработка полученого ответа от камеры(бракуем или нет).
       //Если не бракуем, освобождаем очередь, Если бракуем то взводим бит браковки и освобождаем очередь после снятия сигнала с пушера
       IF "QueueProduct_2".StructQueue[#NumberQueue].ResultRecieved & "QueueProduct_2".StructQueue[#NumberQueue].ResultMeasurementCamera
           & ("QueueProduct_2".StructQueue[#NumberQueue].CurrentImpulseEncodera + "DataBlockHMI".Recipe[0].CountImpTrigerCamera2
           + "DataBlockHMI".Recipe[0].CountImpForRegection2 <= "HWCurrentImpulseEncoder":P) THEN //условия для старта отбраковки

           "AuxaluryBlockProcesseComandeCamera".QuitRejectCam2 := TRUE;
           "DataBlockHMI".AuxilaryBit[1] := TRUE;
           "QueueProduct_2".StructQueue[#NumberQueue].RejectionOn := TRUE;
           "QueueProduct_2".StructQueue[#NumberQueue].ResultRecieved := FALSE;

       ELSIF "QueueProduct_2".StructQueue[#NumberQueue].ResultRecieved & NOT "QueueProduct_2".StructQueue[#NumberQueue].ResultMeasurementCamera THEN

           "QueueProduct_2".StructQueue[#NumberQueue] := "QueueProduct_2".StructQueue[100];

       END_IF;

       //Cнимаем выход отбраковки и скидываем очередь
       IF "QueueProduct_2".StructQueue[#NumberQueue].RejectionOn & ("QueueProduct_2".StructQueue[#NumberQueue].CurrentImpulseEncodera + "DataBlockHMI".Recipe[0].CountImpTrigerCamera2
           + "DataBlockHMI".Recipe[0].CountImpForRegection2 + "DataBlockHMI".Recipe[0].CountImpForResetRegectio1 <= "HWCurrentImpulseEncoder":P) THEN

           "AuxaluryBlockProcesseComandeCamera".QuitRejectCam2 := FALSE;
           "DataBlockHMI".AuxilaryBit[1] := FALSE;
           "QueueProduct_2".StructQueue[#NumberQueue] := "QueueProduct_2".StructQueue[100];

       END_IF;

       IF "DataBlockHMI".Buttons.ButtonWorkRestrictionPusher THEN
           "AuxaluryBlockProcesseComandeCamera".QuitRejectCam2 := FALSE;

       END_IF;


   END_IF;
END_FUNCTION

ORGANIZATION_BLOCK "Main"   // OB1, LAD, ProgramCycle
TITLE = "Main Program Sweep (Cycle)"
{ S7_Optimized_Access := 'TRUE' }
VERSION : 0.1
   VAR_INPUT
      Initial_Call : Bool;   // Initial call of this OB
      Remanence : Bool;   // =True, if remanent data are available
   END_VAR
   VAR_TEMP
      NumberQueue : Int;
   END_VAR
   VAR_TEMP   // added for the SCL form of the ladder/FBD networks
      _w1 : Bool;
      _w2 : Bool;
      _w3 : Bool;
   END_VAR
BEGIN

REGION Network 1: Счетчик отбраковки
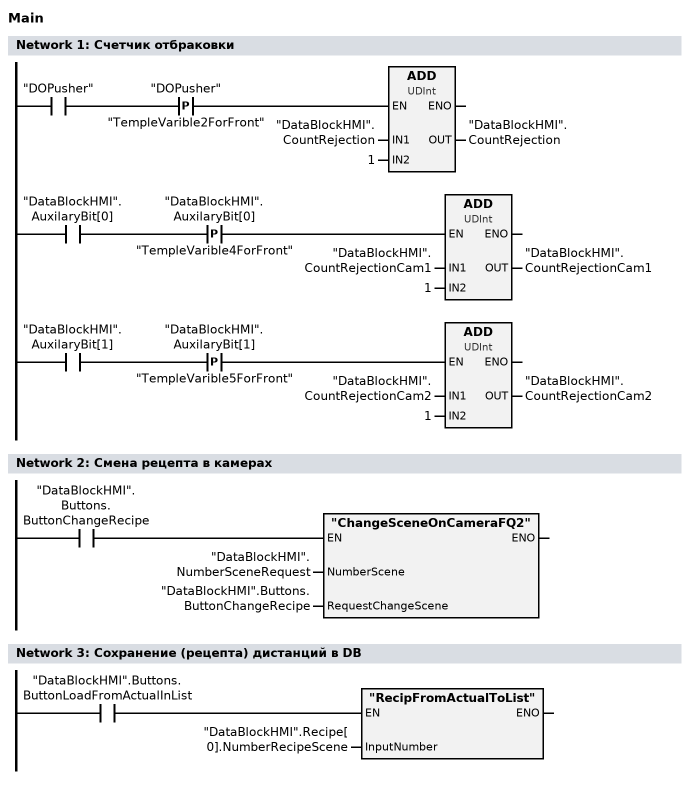
   RUNG wire#powerrail
      Contact( "DOPusher" )
      P_Contact(operand := "DOPusher", bit := "TempleVarible2ForFront")
      { S7_Templates := "SrcType := UDInt" } Add(in1 := "DataBlockHMI".CountRejection, in2 := 1, out => "DataBlockHMI".CountRejection)
   END_RUNG
   RUNG wire#powerrail
      Contact( "DataBlockHMI".AuxilaryBit[0] )
      P_Contact(operand := "DataBlockHMI".AuxilaryBit[0], bit := "TempleVarible4ForFront")
      { S7_Templates := "SrcType := UDInt" } Add(in1 := "DataBlockHMI".CountRejectionCam1, in2 := 1, out => "DataBlockHMI".CountRejectionCam1)
   END_RUNG
   RUNG wire#powerrail
      Contact( "DataBlockHMI".AuxilaryBit[1] )
      P_Contact(operand := "DataBlockHMI".AuxilaryBit[1], bit := "TempleVarible5ForFront")
      { S7_Templates := "SrcType := UDInt" } Add(in1 := "DataBlockHMI".CountRejectionCam2, in2 := 1, out => "DataBlockHMI".CountRejectionCam2)
   END_RUNG
   // the same network as SCL:
   #_w1 := "DOPusher" AND "DOPusher" AND NOT "TempleVarible2ForFront";   // rising edge of "DOPusher"
   "TempleVarible2ForFront" := "DOPusher";
   IF #_w1 THEN "DataBlockHMI".CountRejection := "DataBlockHMI".CountRejection + 1; END_IF;
   #_w2 := "DataBlockHMI".AuxilaryBit[0] AND "DataBlockHMI".AuxilaryBit[0] AND NOT "TempleVarible4ForFront";   // rising edge of "DataBlockHMI".AuxilaryBit[0]
   "TempleVarible4ForFront" := "DataBlockHMI".AuxilaryBit[0];
   IF #_w2 THEN "DataBlockHMI".CountRejectionCam1 := "DataBlockHMI".CountRejectionCam1 + 1; END_IF;
   #_w3 := "DataBlockHMI".AuxilaryBit[1] AND "DataBlockHMI".AuxilaryBit[1] AND NOT "TempleVarible5ForFront";   // rising edge of "DataBlockHMI".AuxilaryBit[1]
   "TempleVarible5ForFront" := "DataBlockHMI".AuxilaryBit[1];
   IF #_w3 THEN "DataBlockHMI".CountRejectionCam2 := "DataBlockHMI".CountRejectionCam2 + 1; END_IF;
END_REGION

REGION Network 2: Смена рецепта в камерах
   RUNG wire#powerrail
      Contact( "DataBlockHMI".Buttons.ButtonChangeRecipe )
      "ChangeSceneOnCameraFQ2"(NumberScene := "DataBlockHMI".NumberSceneRequest, RequestChangeScene := "DataBlockHMI".Buttons.ButtonChangeRecipe)
   END_RUNG
   // the same network as SCL:
   IF "DataBlockHMI".Buttons.ButtonChangeRecipe THEN
       "ChangeSceneOnCameraFQ2"(NumberScene := "DataBlockHMI".NumberSceneRequest,
                               RequestChangeScene := "DataBlockHMI".Buttons.ButtonChangeRecipe);
   END_IF;
END_REGION

REGION Network 3: Сохранение (рецепта) дистанций в DB
   RUNG wire#powerrail
      Contact( "DataBlockHMI".Buttons.ButtonLoadFromActualInList )
      "RecipFromActualToList"(InputNumber := "DataBlockHMI".Recipe[0].NumberRecipeScene)
   END_RUNG
   // the same network as SCL:
   IF "DataBlockHMI".Buttons.ButtonLoadFromActualInList THEN
       "RecipFromActualToList"(InputNumber := "DataBlockHMI".Recipe[0].NumberRecipeScene);
   END_IF;
END_REGION
END_ORGANIZATION_BLOCK

ORGANIZATION_BLOCK "ProcessingQueue"   // OB30, LAD, CyclicInterrupt
{ S7_Optimized_Access := 'TRUE' }
VERSION : 0.1
// В этом блоке читаем с камер, обрабатываем очереди, и записываем в камеры
   VAR_INPUT
      Initial_Call : Bool;   // Initial call of this OB
      Event_Count : Int;   // Events discarded
   END_VAR
   VAR_TEMP
      NumberQueue : Int;
      NumberQueue2 : Int;
   END_VAR
BEGIN

REGION Network 1 (SCL): Чтение с камер
   //Чтение с первой камеры

   POKE_BLK(area_src := 16#81,
            dbNumber_src := 0,
            byteOffset_src := 68,
            area_dest := 16#84,
            dbNumber_dest := 2,
            byteOffset_dest := 0,
            count := 144);

   //Чтение со 2ой камеры
   POKE_BLK(area_src := 16#81,
            dbNumber_src := 0,
            byteOffset_src := 212,
            area_dest := 16#84,
            dbNumber_dest := 2,
            byteOffset_dest := 164,
            count := 144);
END_REGION

REGION Network 2 (SCL)
   // Обработак очериди продкута камерой
   IF "InputOutputCamer".InputFromCamera1.RUN OR "InputOutputCamer".InputFromCamera2.RUN THEN
       FOR #NumberQueue := 0 TO 20 DO
           IF NOT "DataBlockHMI".Buttons.ButtonWorkOffCam1 THEN
               "ProcessingQueue1"(#NumberQueue);
           END_IF;
           IF NOT "DataBlockHMI".Buttons.ButtonWorkOffCam2 THEN
               "ProcessingQueue2"(#NumberQueue);

           END_IF;
       END_FOR;
   END_IF;
END_REGION

REGION Network 3 (SCL): Запись в камеры
   //Запись в первую камеру
   POKE_BLK(area_src := 16#84,
            dbNumber_src := 2,
            byteOffset_src := 144,
            area_dest := 16#82,
            dbNumber_dest := 0,
            byteOffset_dest := 2,
            count := 20);
   //Запись во вторую камеру
   POKE_BLK(area_src := 16#84,
            dbNumber_src := 2,
            byteOffset_src := 308,
            area_dest := 16#82,
            dbNumber_dest := 0,
            byteOffset_dest := 22,
            count := 20);
END_REGION

REGION Network 4: Работа пушера
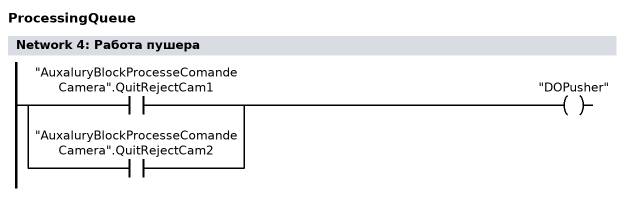
   RUNG wire#powerrail
      Contact( "AuxaluryBlockProcesseComandeCamera".QuitRejectCam1 )
      wire#w1
      Coil( "DOPusher" )
   END_RUNG
   RUNG wire#powerrail
      Contact( "AuxaluryBlockProcesseComandeCamera".QuitRejectCam2 )
   END_RUNG wire#w1
   // the same network as SCL:
   "DOPusher" := "AuxaluryBlockProcesseComandeCamera".QuitRejectCam1 OR "AuxaluryBlockProcesseComandeCamera".QuitRejectCam2;
END_REGION
END_ORGANIZATION_BLOCK

ORGANIZATION_BLOCK "Hardware interrupt"   // OB40, LAD, HWProcessInterrupt
{ S7_Optimized_Access := 'TRUE' }
VERSION : 0.1
   VAR_INPUT
      LADDR : Hw_Io;   // Hardware identifier
      USI : Word;   // User structure identifier
      IChannel : USInt;   // Interrupt channel number
      EventType : Byte;   // EventType
   END_VAR
BEGIN

REGION Network 1
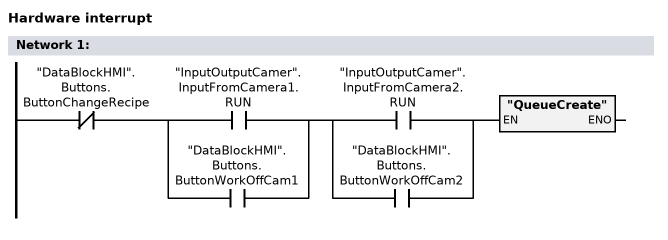
   RUNG wire#powerrail
      I_Contact( "DataBlockHMI".Buttons.ButtonChangeRecipe )
      wire#w1
      Contact( "InputOutputCamer".InputFromCamera1.RUN )
      wire#w2
      Contact( "InputOutputCamer".InputFromCamera2.RUN )
      wire#w3
      "QueueCreate"()
   END_RUNG
   RUNG wire#w1
      Contact( "DataBlockHMI".Buttons.ButtonWorkOffCam1 )
   END_RUNG wire#w2
   RUNG wire#w2
      Contact( "DataBlockHMI".Buttons.ButtonWorkOffCam2 )
   END_RUNG wire#w3
   // the same network as SCL:
   IF NOT "DataBlockHMI".Buttons.ButtonChangeRecipe AND ("InputOutputCamer".InputFromCamera1.RUN OR "DataBlockHMI".Buttons.ButtonWorkOffCam1) AND ("InputOutputCamer".InputFromCamera2.RUN OR "DataBlockHMI".Buttons.ButtonWorkOffCam2) THEN
       "QueueCreate"();
   END_IF;
END_REGION
END_ORGANIZATION_BLOCK